// TIA Portal V20 export
// export: Created 2026-10-12T05:42:32.5058003Z, ExportSetting WithDefaults, DisplayName Totally Integrated Automation Portal, DisplayVersion V20, DisplayName TIA Portal Openness, DisplayVersion V20, DisplayName TIA Portal Teamcenter Gateway, DisplayVersion V20, DisplayName TIA Portal Version Control Interface, DisplayVersion V20, DisplayName SINAMICS Startdrive Advanced, DisplayVersion V20 SP1 Update 2, DisplayName SINAMICS Startdrive G110M, G120, G120C, G120D, G120P, G115D, DisplayVersion V20 SP1 Update 2, DisplayName SINAMICS Startdrive G130, G150, S120, S150, SINAMICS MV, G220, S200, S210, DisplayVersion V20 SP1 Update 2, DisplayName STEP 7 Professional, DisplayVersion V20, DisplayName STEP 7 Safety, DisplayVersion V20, DisplayName WinCC Basic/Comfort/Advanced, DisplayVersion V20, DisplayName WinCC Professional, DisplayVersion V20, DisplayName WinCC Unified, DisplayVersion V20
FUNCTION "FRK_SeqBegin" : Void   // FC124, SCL
{ S7_Optimized_Access := 'TRUE' }
VERSION : 0.1
// Shared sequence services. The examples generator binds Core enum constants.
// stored: AutoNumber true, IsIECCheckEnabled false, SetENOAutomatically false, UDAEnableTagReadback false
   VAR_INPUT
      Run : Bool;
      Reset : Bool;
      OwnerIndex : DInt;
      ChainIndex : DInt;
      BranchIndex : DInt;
      Delta : Time;
   END_VAR
   VAR_IN_OUT
      Seq : "FRK_SequenceCtx";
   END_VAR
BEGIN

   #Seq.Scan := #Seq.Scan + 1;
   #Seq.Restart := #Reset OR (#Run AND NOT #Seq.RunPrevious);
   #Seq.RunPrevious := #Run;
   #Seq.OwnerIndex := #OwnerIndex;
   #Seq.ChainIndex := #ChainIndex;
   #Seq.BranchIndex := #BranchIndex;
   #Seq.RetVal := 0;
   #Seq.Pending := FALSE;
   #Seq.CommandFailed := FALSE;
   #Seq.CommandIssued := FALSE;
   #Seq.Awaiting := '';
   IF NOT #Run OR #Seq.Restart THEN
       #Seq.Step := 0;
       #Seq.RecordedStep := -1;
       #Seq.Visit := #Seq.Visit + 1;
       #Seq.Done := FALSE;
       #Seq.Error := FALSE;
       #Seq.StartLatched := FALSE;
       #Seq.Elapsed := T#0ms;
       #Seq.DelayElapsed := T#0ms;
       #Seq.ErrorDiagnostic.ReasonCode := 0;
   END_IF;
   #Seq.Running := #Run AND NOT #Seq.Done AND NOT #Seq.Error
   AND #OwnerIndex > 0 AND #ChainIndex > 0;
   #Seq.ScanStep := #Seq.Step;
   IF #Seq.Running AND #Delta > T#0ms THEN
       #Seq.Elapsed := #Seq.Elapsed + #Delta;
   END_IF;
END_FUNCTION
